(* IEC 61131-3 sources: plc-iiot-stack/src/POUs/Json/FB_JsonBuilder, 21 files *)

(* ---- FB_JsonBuilder.decl.st ---- *)
// Назначение: построитель плоского объекта JSON в буфере STRING(GVL_Const.MQTT_PAYLOAD_LEN) побайтно, без
//             CONCAT (стандартные строковые функции ограничены 255 символами). Ключи и строки
//             экранируются, REAL — с фиксированным числом знаков без хвостовых нулей, NaN и
//             бесконечность — null, целые — LINT. Переполнение буфера фиксируется флагом xOverflow:
//             неполный JSON публиковать нельзя.
//             Порядок: Begin(), Add...() для каждого поля, Finish() (TRUE — объект закончен и помещается).
// Автор:      kr0nsch
// Версия:     0.1.0
// Документ:   docs/plc_mqtt.md, раздел «Построение JSON»
FUNCTION_BLOCK FB_JsonBuilder
VAR_OUTPUT
    sJson : STRING(GVL_Const.MQTT_PAYLOAD_LEN);   // текст JSON
    uiLen : UINT;                                  // длина текста, байт
    xOverflow : BOOL;                              // буфер переполнен: текст неполный
END_VAR
VAR
    xNeedComma : BOOL;                             // перед следующим полем нужна запятая
END_VAR

(* ---- AddBool.method.decl.st ---- *)
// Поле true или false.
METHOD AddBool
VAR_INPUT
    sKey : STRING(GVL_Const.JSON_KEY_LEN);
    xValue : BOOL;
END_VAR

(* ---- AddBool.method.impl.st ---- *)
AppendKey(sKeyName := sKey);
IF xValue THEN
    AppendRaw(sText := 'true');
ELSE
    AppendRaw(sText := 'false');
END_IF

(* ---- AddInt.method.decl.st ---- *)
// Поле с целым числом (любой целый тип приводится к LINT).
METHOD AddInt
VAR_INPUT
    sKey : STRING(GVL_Const.JSON_KEY_LEN);
    liValue : LINT;
END_VAR

(* ---- AddNull.method.decl.st ---- *)
// Поле со значением null.
METHOD AddNull
VAR_INPUT
    sKey : STRING(GVL_Const.JSON_KEY_LEN);
END_VAR

(* ---- AddReal.method.decl.st ---- *)
// Поле с числом: uiDecimals знаков после точки (не больше JSON_REAL_DECIMALS_MAX), хвостовые нули
// отбрасываются; NaN, бесконечность и слишком большие числа — null. REAL приводится к LREAL.
METHOD AddReal
VAR_INPUT
    sKey : STRING(GVL_Const.JSON_KEY_LEN);
    lrValue : LREAL;
    uiDecimals : UINT;
END_VAR

(* ---- AddString.method.decl.st ---- *)
// Поле со строковым значением; кавычки, обратная косая черта и управляющие символы экранируются.
METHOD AddString
VAR_INPUT
    sKey : STRING(GVL_Const.JSON_KEY_LEN);
    sValue : STRING(GVL_Const.JSON_STR_LEN);
END_VAR

(* ---- AppendByte.method.decl.st ---- *)
// Дописать один байт; места нет — xOverflow, буфер не меняется.
METHOD PRIVATE AppendByte
VAR_INPUT
    bChar : BYTE;
END_VAR

(* ---- AppendByte.method.impl.st ---- *)
IF uiLen >= GVL_Const.MQTT_PAYLOAD_LEN THEN
    xOverflow := TRUE;
    RETURN;
END_IF
sJson[uiLen] := bChar;
uiLen := uiLen + 1;
sJson[uiLen] := GVL_Const.ASCII_NUL;

(* ---- AppendEscaped.method.decl.st ---- *)
// Дописать строку с экранированием JSON: \" \\ \n \r \t \b \f; прочие управляющие символы и байты
// не из ASCII — \u00XX (байт как символ Latin-1; строки ПЛК в этом проекте — ASCII).
METHOD PRIVATE AppendEscaped
VAR_INPUT
    sText : STRING(GVL_Const.JSON_STR_LEN);
END_VAR
VAR
    uiTextLen : UINT;
    uiIdx : UINT;
    bCh : BYTE;
END_VAR

(* ---- AppendEscaped.method.impl.st ---- *)
uiTextLen := INT_TO_UINT(LEN(sText));
uiIdx := 0;
WHILE uiIdx < uiTextLen DO
    bCh := sText[uiIdx];
    IF bCh = GVL_Const.ASCII_QUOTE OR bCh = GVL_Const.ASCII_BACKSLASH THEN
        AppendByte(bChar := GVL_Const.ASCII_BACKSLASH);
        AppendByte(bChar := bCh);
    ELSIF bCh = GVL_Const.ASCII_LF THEN
        AppendByte(bChar := GVL_Const.ASCII_BACKSLASH);
        AppendByte(bChar := GVL_Const.ASCII_LOWER_N);
    ELSIF bCh = GVL_Const.ASCII_CR THEN
        AppendByte(bChar := GVL_Const.ASCII_BACKSLASH);
        AppendByte(bChar := GVL_Const.ASCII_LOWER_R);
    ELSIF bCh = GVL_Const.ASCII_TAB THEN
        AppendByte(bChar := GVL_Const.ASCII_BACKSLASH);
        AppendByte(bChar := GVL_Const.ASCII_LOWER_T);
    ELSIF bCh = GVL_Const.ASCII_BS THEN
        AppendByte(bChar := GVL_Const.ASCII_BACKSLASH);
        AppendByte(bChar := GVL_Const.ASCII_LOWER_B);
    ELSIF bCh = GVL_Const.ASCII_FF THEN
        AppendByte(bChar := GVL_Const.ASCII_BACKSLASH);
        AppendByte(bChar := GVL_Const.ASCII_LOWER_F);
    ELSIF bCh <= GVL_Const.ASCII_CTRL_LAST OR bCh > GVL_Const.ASCII_LAST THEN
        AppendByte(bChar := GVL_Const.ASCII_BACKSLASH);
        AppendByte(bChar := GVL_Const.ASCII_LOWER_U);
        AppendByte(bChar := GVL_Const.ASCII_ZERO);
        AppendByte(bChar := GVL_Const.ASCII_ZERO);
        AppendHexDigit(bNibble := SHR(bCh, GVL_Const.NIBBLE_BITS));
        AppendHexDigit(bNibble := bCh AND GVL_Const.NIBBLE_MASK);
    ELSE
        AppendByte(bChar := bCh);
    END_IF
    uiIdx := uiIdx + 1;
END_WHILE

(* ---- AppendHexDigit.method.decl.st ---- *)
// Дописать шестнадцатеричную цифру 0..f (младшие 4 бита bNibble).
METHOD PRIVATE AppendHexDigit
VAR_INPUT
    bNibble : BYTE;
END_VAR
VAR
    bDigit : BYTE;
END_VAR

(* ---- AppendHexDigit.method.impl.st ---- *)
bDigit := bNibble AND GVL_Const.NIBBLE_MASK;
IF bDigit < GVL_Const.HEX_LETTER_START THEN
    AppendByte(bChar := GVL_Const.ASCII_ZERO + bDigit);
ELSE
    AppendByte(bChar := GVL_Const.ASCII_LOWER_A + (bDigit - GVL_Const.HEX_LETTER_START));
END_IF

(* ---- AppendInt.method.decl.st ---- *)
// Дописать десятичную запись целого со знаком (включая минимальное значение LINT).
METHOD PRIVATE AppendInt
VAR_INPUT
    liNumber : LINT;
END_VAR
VAR
    uliMagnitude : ULINT;
END_VAR

(* ---- AppendInt.method.impl.st ---- *)
IF liNumber < 0 THEN
    AppendByte(bChar := GVL_Const.ASCII_MINUS);
    // -(x + 1) не переполняется и для минимального LINT
    uliMagnitude := LINT_TO_ULINT(-(liNumber + 1)) + 1;
ELSE
    uliMagnitude := LINT_TO_ULINT(liNumber);
END_IF
AppendUlint(uliNumber := uliMagnitude);

(* ---- AppendKey.method.decl.st ---- *)
// Запятая (если поле не первое), ключ в кавычках и двоеточие.
METHOD PRIVATE AppendKey
VAR_INPUT
    sKeyName : STRING(GVL_Const.JSON_KEY_LEN);
END_VAR

(* ---- AppendKey.method.impl.st ---- *)
IF xNeedComma THEN
    AppendByte(bChar := GVL_Const.ASCII_COMMA);
END_IF
xNeedComma := TRUE;
AppendByte(bChar := GVL_Const.ASCII_QUOTE);
AppendEscaped(sText := sKeyName);
AppendByte(bChar := GVL_Const.ASCII_QUOTE);
AppendByte(bChar := GVL_Const.ASCII_COLON);

(* ---- AppendRaw.method.decl.st ---- *)
// Дописать текст как есть (литералы JSON, цифры).
METHOD PRIVATE AppendRaw
VAR_INPUT
    sText : STRING(GVL_Const.JSON_STR_LEN);
END_VAR
VAR
    uiTextLen : UINT;
    uiIdx : UINT;
END_VAR

(* ---- AppendReal.method.decl.st ---- *)
// Дописать число с uiDecimalsMax знаками (округление до ближайшего), без хвостовых нулей; -0 пишется как 0.
METHOD PRIVATE AppendReal
VAR_INPUT
    lrNumber : LREAL;
    uiDecimalsMax : UINT;
END_VAR
VAR
    uiDecimals : UINT;
    uiIdx : UINT;
    uliScale : ULINT;          // 10^uiDecimals
    lrScaled : LREAL;
    uliScaled : ULINT;
    uliFrac : ULINT;
    uiFracDigits : UINT;       // значащих знаков дробной части после отбрасывания нулей
    uiDigits : UINT;
    uliTmp : ULINT;
END_VAR

(* ---- AppendReal.method.impl.st ---- *)
IF NOT F_IsFiniteLreal(lrValue := lrNumber) THEN
    AppendRaw(sText := 'null');
    RETURN;
END_IF
uiDecimals := MIN(uiDecimalsMax, GVL_Const.JSON_REAL_DECIMALS_MAX);
uliScale := 1;
FOR uiIdx := 1 TO uiDecimals DO
    uliScale := uliScale * GVL_Const.DECIMAL_BASE;
END_FOR
lrScaled := ABS(lrNumber) * ULINT_TO_LREAL(uliScale);
IF lrScaled >= GVL_Const.JSON_NUM_SCALED_MAX THEN
    AppendRaw(sText := 'null');
    RETURN;
END_IF
// преобразование LREAL -> ULINT в CODESYS округляет до ближайшего целого
uliScaled := LREAL_TO_ULINT(lrScaled);
IF lrNumber < 0.0 AND uliScaled > 0 THEN
    AppendByte(bChar := GVL_Const.ASCII_MINUS);
END_IF
AppendUlint(uliNumber := uliScaled / uliScale);
uliFrac := uliScaled MOD uliScale;
IF uliFrac > 0 THEN
    AppendByte(bChar := GVL_Const.ASCII_DOT);
    uiFracDigits := uiDecimals;
    WHILE (uliFrac MOD GVL_Const.DECIMAL_BASE) = 0 DO
        uliFrac := uliFrac / GVL_Const.DECIMAL_BASE;
        uiFracDigits := uiFracDigits - 1;
    END_WHILE
    // ведущие нули дробной части: значащих цифр у остатка меньше, чем знаков
    uliTmp := uliFrac;
    uiDigits := 0;
    WHILE uliTmp > 0 DO
        uliTmp := uliTmp / GVL_Const.DECIMAL_BASE;
        uiDigits := uiDigits + 1;
    END_WHILE
    WHILE uiDigits < uiFracDigits DO
        AppendByte(bChar := GVL_Const.ASCII_ZERO);
        uiDigits := uiDigits + 1;
    END_WHILE
    AppendUlint(uliNumber := uliFrac);
END_IF

(* ---- AppendUlint.method.decl.st ---- *)
// Дописать десятичную запись целого без знака.
METHOD PRIVATE AppendUlint
VAR_INPUT
    uliNumber : ULINT;
END_VAR
VAR
    aDigits : ARRAY[0..GVL_Const.ULINT_DIGITS_MAX - 1] OF BYTE;   // цифры с младшей
    uiCount : UINT;
    uliRest : ULINT;
END_VAR
